Staubli VAL3: sPointTemplate.pjx

--- sPointTemplate.pjx ---
Parameters version=s8.10.3Cs9_BS2093 stackSize=5000 millimeterUnit=true
Program file=start.pgx
Program file=stop.pgx
Data file=sPointTemplate.dtx

--- sPointTemplate.dtx ---
public bool bActive
public pointRx pPointRx = {fatherId=world[0]}
public string sName

--- start.pgx ---
program start()
begin
end

--- stop.pgx ---
program stop()
begin
end
